Fanuc KAREL source: kb00160.KL

PROGRAM KB00160
%NOLOCKGROUP
VAR
P1 : FILE
P2:INTEGER
P3:INTEGER
P4:INTEGER
BEGIN
P2=1
P3=1
P4=1
SET_CURSOR(P1,P2,P3,P4)
END KB00160
